Fanuc KAREL source: kb00022.KL

-- PROVISIONAL review KL for V1013-1; original PC SHA256 7e2d2f0999714e962cbe4562b6e2f806b2ce2e05d8a9eaebfc6cdf05dc343751
-- Incomplete behavior may be omitted. Consult companion uncertainty JSON. Do not deploy.
PROGRAM KB00022
%NOLOCKGROUP
BEGIN
  -- UNRESOLVED_PC offsets 5-12; opcodes 9D,23
  -- UNRESOLVED_PC offsets 17-27; opcodes 27,22,31
  -- UNRESOLVED_PC offsets 32-36; opcodes 7F
END KB00022
